(* IEC 61131-3 sources: trust-platform/examples/OSCAT/hvac_air_handling_unit/oop/src, 3 files *)

(* ---- Main.st ---- *)
(* Pattern role: IAhuStrategy is the contract boundary for the Strategy example. *)
INTERFACE IAhuStrategy EXTENDS IComponent
    PROPERTY ModeId : INT
    GET
    END_GET
    END_PROPERTY

    PROPERTY Output : REAL
    GET
    END_GET
    END_PROPERTY

    METHOD AcceptsCommand : BOOL
    VAR_INPUT
        SmokeClear : BOOL;
        FreezeStatClear : BOOL;
    END_VAR
    END_METHOD

    METHOD Update : REAL
    VAR_INPUT
        SupplyTemp : REAL;
        ScheduledSetpoint : REAL;
        OutdoorTemp : REAL;
    END_VAR
    END_METHOD
END_INTERFACE

(* Pattern role: EcoStrategy is a concrete implementation in the Strategy example. *)
FUNCTION_BLOCK EcoStrategy IMPLEMENTS IAhuStrategy
VAR
    ReadyValue : BOOL;
    ErrorValue : BOOL;
    ErrorIdValue : WORD;
    StatusValue : BYTE;
    OutputValue : REAL;
    Filter : Pt1Filter;
END_VAR

METHOD PUBLIC Initialize
ReadyValue := TRUE;
Filter.Initialize();
Filter.Configure(TimeConstant := T#5s, Gain := REAL#1.0);
ClearError();
END_METHOD

METHOD PUBLIC Reset
OutputValue := REAL#0.0;
ClearError();
END_METHOD

METHOD PUBLIC ClearError
ErrorValue := FALSE;
ErrorIdValue := WORD#0;
StatusValue := BYTE#0;
END_METHOD

METHOD PUBLIC Snapshot : ComponentStatus
VAR
    Result : ComponentStatus;
END_VAR
Result.Ready := ReadyValue;
Result.Error := ErrorValue;
Result.ErrorId := ErrorIdValue;
Result.Status := StatusValue;
Snapshot := Result;
END_METHOD

METHOD PUBLIC AcceptsCommand : BOOL
VAR_INPUT
    SmokeClear : BOOL;
    FreezeStatClear : BOOL;
END_VAR
AcceptsCommand := SmokeClear AND FreezeStatClear;
END_METHOD

METHOD PUBLIC Update : REAL
VAR_INPUT
    SupplyTemp : REAL;
    ScheduledSetpoint : REAL;
    OutdoorTemp : REAL;
END_VAR
VAR
    Error : REAL;
END_VAR
(* Filter is kept on the snapshot side for telemetry smoothing; the
   deadband and gain operate on the raw supply temp so the controller
   reacts to step changes within the same scan. *)
Filter.Update(Sample := SupplyTemp);
Error := ScheduledSetpoint - SupplyTemp;
IF ABS(Error) <= REAL#2.0 THEN
    OutputValue := REAL#0.0;
ELSE
    OutputValue := LIMIT(REAL#0.0, Error * REAL#8.0, REAL#100.0);
END_IF;
Update := OutputValue;
END_METHOD

PUBLIC PROPERTY ModeId : INT
GET
    ModeId := INT#1;
END_GET
END_PROPERTY

PUBLIC PROPERTY Output : REAL
GET
    Output := OutputValue;
END_GET
END_PROPERTY

PUBLIC PROPERTY Ready : BOOL
GET
    Ready := ReadyValue;
END_GET
END_PROPERTY

PUBLIC PROPERTY Error : BOOL
GET
    Error := ErrorValue;
END_GET
END_PROPERTY

PUBLIC PROPERTY ErrorId : WORD
GET
    ErrorId := ErrorIdValue;
END_GET
END_PROPERTY

PUBLIC PROPERTY Status : BYTE
GET
    Status := StatusValue;
END_GET
END_PROPERTY
END_FUNCTION_BLOCK

(* Pattern role: ComfortStrategy is a concrete implementation in the Strategy example. *)
FUNCTION_BLOCK ComfortStrategy IMPLEMENTS IAhuStrategy
VAR
    ReadyValue : BOOL;
    ErrorValue : BOOL;
    ErrorIdValue : WORD;
    StatusValue : BYTE;
    OutputValue : REAL;
    Filter : Pt1Filter;
END_VAR

METHOD PUBLIC Initialize
ReadyValue := TRUE;
Filter.Initialize();
Filter.Configure(TimeConstant := T#1s, Gain := REAL#1.0);
ClearError();
END_METHOD

METHOD PUBLIC Reset
OutputValue := REAL#0.0;
ClearError();
END_METHOD

METHOD PUBLIC ClearError
ErrorValue := FALSE;
ErrorIdValue := WORD#0;
StatusValue := BYTE#0;
END_METHOD

METHOD PUBLIC Snapshot : ComponentStatus
VAR
    Result : ComponentStatus;
END_VAR
Result.Ready := ReadyValue;
Result.Error := ErrorValue;
Result.ErrorId := ErrorIdValue;
Result.Status := StatusValue;
Snapshot := Result;
END_METHOD

METHOD PUBLIC AcceptsCommand : BOOL
VAR_INPUT
    SmokeClear : BOOL;
    FreezeStatClear : BOOL;
END_VAR
AcceptsCommand := SmokeClear;
END_METHOD

METHOD PUBLIC Update : REAL
VAR_INPUT
    SupplyTemp : REAL;
    ScheduledSetpoint : REAL;
    OutdoorTemp : REAL;
END_VAR
VAR
    Error : REAL;
END_VAR
(* Same approach as Eco: deadband/gain on raw supply, filter
   advanced for telemetry only. Strict inequality so Comfort reacts
   at the deadband boundary (tighter response than Eco). *)
Filter.Update(Sample := SupplyTemp);
Error := ScheduledSetpoint - SupplyTemp;
IF ABS(Error) < REAL#0.5 THEN
    OutputValue := REAL#0.0;
ELSE
    OutputValue := LIMIT(REAL#0.0, Error * REAL#20.0, REAL#100.0);
END_IF;
Update := OutputValue;
END_METHOD

PUBLIC PROPERTY ModeId : INT
GET
    ModeId := INT#2;
END_GET
END_PROPERTY

PUBLIC PROPERTY Output : REAL
GET
    Output := OutputValue;
END_GET
END_PROPERTY

PUBLIC PROPERTY Ready : BOOL
GET
    Ready := ReadyValue;
END_GET
END_PROPERTY

PUBLIC PROPERTY Error : BOOL
GET
    Error := ErrorValue;
END_GET
END_PROPERTY

PUBLIC PROPERTY ErrorId : WORD
GET
    ErrorId := ErrorIdValue;
END_GET
END_PROPERTY

PUBLIC PROPERTY Status : BYTE
GET
    Status := StatusValue;
END_GET
END_PROPERTY
END_FUNCTION_BLOCK

(* Pattern role: FrostProtectStrategy is a concrete implementation in the Strategy example. *)
FUNCTION_BLOCK FrostProtectStrategy IMPLEMENTS IAhuStrategy
VAR
    ReadyValue : BOOL;
    ErrorValue : BOOL;
    ErrorIdValue : WORD;
    StatusValue : BYTE;
    OutputValue : REAL;
END_VAR

METHOD PUBLIC Initialize
ReadyValue := TRUE;
ClearError();
END_METHOD

METHOD PUBLIC Reset
OutputValue := REAL#0.0;
ClearError();
END_METHOD

METHOD PUBLIC ClearError
ErrorValue := FALSE;
ErrorIdValue := WORD#0;
StatusValue := BYTE#0;
END_METHOD

METHOD PUBLIC Snapshot : ComponentStatus
VAR
    Result : ComponentStatus;
END_VAR
Result.Ready := ReadyValue;
Result.Error := ErrorValue;
Result.ErrorId := ErrorIdValue;
Result.Status := StatusValue;
Snapshot := Result;
END_METHOD

METHOD PUBLIC AcceptsCommand : BOOL
VAR_INPUT
    SmokeClear : BOOL;
    FreezeStatClear : BOOL;
END_VAR
AcceptsCommand := SmokeClear;
END_METHOD

METHOD PUBLIC Update : REAL
VAR_INPUT
    SupplyTemp : REAL;
    ScheduledSetpoint : REAL;
    OutdoorTemp : REAL;
END_VAR
VAR
    FrostTarget : REAL;
END_VAR
FrostTarget := MAX(ScheduledSetpoint, REAL#5.0);
OutputValue := LIMIT(REAL#20.0, (FrostTarget - SupplyTemp) * REAL#30.0, REAL#100.0);
Update := OutputValue;
END_METHOD

PUBLIC PROPERTY ModeId : INT
GET
    ModeId := INT#3;
END_GET
END_PROPERTY

PUBLIC PROPERTY Output : REAL
GET
    Output := OutputValue;
END_GET
END_PROPERTY

PUBLIC PROPERTY Ready : BOOL
GET
    Ready := ReadyValue;
END_GET
END_PROPERTY

PUBLIC PROPERTY Error : BOOL
GET
    Error := ErrorValue;
END_GET
END_PROPERTY

PUBLIC PROPERTY ErrorId : WORD
GET
    ErrorId := ErrorIdValue;
END_GET
END_PROPERTY

PUBLIC PROPERTY Status : BYTE
GET
    Status := StatusValue;
END_GET
END_PROPERTY
END_FUNCTION_BLOCK

(* Composition role: AhuController owns the collaborating objects used by this Strategy example. *)
FUNCTION_BLOCK AhuController
VAR
    Eco : EcoStrategy;
    Comfort : ComfortStrategy;
    Frost : FrostProtectStrategy;
    ActiveStrategy : IAhuStrategy;
    StateValue : INT;
    ActiveModeValue : INT;
    HeatingCommandValue : REAL;
    AlarmActiveValue : BOOL;
    AlarmCodeValue : DWORD;
    RuntimeFan : OntimeMeter;
    AlarmQueue : DwordFifo16;
END_VAR

METHOD PUBLIC Initialize
Eco.Initialize();
Comfort.Initialize();
Frost.Initialize();
RuntimeFan.Initialize();
RuntimeFan.Reset();
AlarmQueue.Initialize();
AlarmQueue.Reset();
StateValue := INT#0;
ActiveModeValue := INT#0;
HeatingCommandValue := REAL#0.0;
AlarmActiveValue := FALSE;
AlarmCodeValue := DWORD#0;
END_METHOD

METHOD PRIVATE RaiseAlarm
VAR_INPUT
    Code : DWORD;
END_VAR
AlarmActiveValue := TRUE;
AlarmCodeValue := Code;
StateValue := INT#900;
IF AlarmQueue.Push(Value := Code) THEN
END_IF;
END_METHOD

METHOD PUBLIC Update : REAL
VAR_INPUT
    ModeRequest : INT;
    OutdoorTemp : REAL;
    SupplyTemp : REAL;
    SupplySetpoint : REAL;
    SmokeClear : BOOL;
    FreezeStatClear : BOOL;
    SupplyFanHealthy : BOOL;
END_VAR
IF NOT SmokeClear THEN
    RaiseAlarm(Code := DWORD#16#A100);
    HeatingCommandValue := REAL#0.0;
ELSE
    IF (OutdoorTemp < REAL#-5.0) OR NOT FreezeStatClear THEN
        ActiveStrategy := Frost;
    ELSIF ModeRequest = INT#1 THEN
        ActiveStrategy := Eco;
    ELSE
        ActiveStrategy := Comfort;
    END_IF;

    ActiveModeValue := ActiveStrategy.ModeId;
    IF NOT SupplyFanHealthy THEN
        RaiseAlarm(Code := DWORD#16#A101);
    ELSIF ActiveStrategy.AcceptsCommand(SmokeClear := SmokeClear, FreezeStatClear := FreezeStatClear) THEN
        StateValue := INT#200;
        HeatingCommandValue := ActiveStrategy.Update(SupplyTemp := SupplyTemp, ScheduledSetpoint := SupplySetpoint, OutdoorTemp := OutdoorTemp);
        RuntimeFan.Update(Input := TRUE);
    ELSE
        RaiseAlarm(Code := DWORD#16#B100);
    END_IF;
END_IF;
Update := HeatingCommandValue;
END_METHOD

PUBLIC PROPERTY State : INT
GET
    State := StateValue;
END_GET
END_PROPERTY

PUBLIC PROPERTY ActiveMode : INT
GET
    ActiveMode := ActiveModeValue;
END_GET
END_PROPERTY

PUBLIC PROPERTY HeatingCommand : REAL
GET
    HeatingCommand := HeatingCommandValue;
END_GET
END_PROPERTY

PUBLIC PROPERTY AlarmActive : BOOL
GET
    AlarmActive := AlarmActiveValue;
END_GET
END_PROPERTY
END_FUNCTION_BLOCK

(* Scan role: Main wires the example objects and exposes the PLC call path under test. *)
PROGRAM Main
VAR
    Ahu : AhuController;
    Initialized : BOOL;
    ModeRequest : INT;
    OutdoorTempRaw : INT;
    SupplyTempRaw : INT;
    SmokeClear : BOOL;
    FreezeStatClear : BOOL;
    SupplyFanHealthy : BOOL;
    HeatingValveRaw : INT;
    SupplyFanEnable : BOOL;
    FireAlarmRelay : BOOL;
    OutdoorTemp : REAL;
    SupplyTemp : REAL;
END_VAR

OutdoorTemp := TO_REAL(OutdoorTempRaw) / REAL#10.0;
SupplyTemp := TO_REAL(SupplyTempRaw) / REAL#10.0;
(* Initialize once on cold start; scanning Initialize every cycle would
   reset RuntimeFan, clear AlarmQueue, and force StateValue back to 0. *)
IF NOT Initialized THEN
    Ahu.Initialize();
    Initialized := TRUE;
END_IF;
HeatingValveRaw := TO_INT(Ahu.Update(ModeRequest := ModeRequest, OutdoorTemp := OutdoorTemp, SupplyTemp := SupplyTemp, SupplySetpoint := REAL#21.0, SmokeClear := SmokeClear, FreezeStatClear := FreezeStatClear, SupplyFanHealthy := SupplyFanHealthy) * REAL#10.0);
SupplyFanEnable := NOT Ahu.AlarmActive;
FireAlarmRelay := NOT SmokeClear;
END_PROGRAM

(* ---- Configuration.st ---- *)
CONFIGURATION AhuOopConfiguration
RESOURCE AhuOop ON PLC
    TASK MainTask (INTERVAL := T#100ms, PRIORITY := 1);
    PROGRAM Ahu WITH MainTask : Main;
END_RESOURCE
VAR_CONFIG
    Ahu.ModeRequest AT %IW0 : INT;
    Ahu.OutdoorTempRaw AT %IW2 : INT;
    Ahu.SupplyTempRaw AT %IW4 : INT;
    Ahu.SmokeClear AT %IX0.0 : BOOL;
    Ahu.FreezeStatClear AT %IX0.1 : BOOL;
    Ahu.SupplyFanHealthy AT %IX0.2 : BOOL;
    Ahu.HeatingValveRaw AT %QW0 : INT;
    Ahu.SupplyFanEnable AT %QX0.0 : BOOL;
    Ahu.FireAlarmRelay AT %QX0.1 : BOOL;
END_VAR
END_CONFIGURATION

(* ---- Tests.st ---- *)
TEST_PROGRAM AhuStrategySelectsModeSpecificObjects
VAR
    Ahu : AhuController;
    EcoCommand : REAL;
    ComfortCommand : REAL;
    FrostCommand : REAL;
END_VAR

Ahu.Initialize();
EcoCommand := Ahu.Update(ModeRequest := INT#1, OutdoorTemp := REAL#10.0, SupplyTemp := REAL#18.0, SupplySetpoint := REAL#21.0, SmokeClear := TRUE, FreezeStatClear := TRUE, SupplyFanHealthy := TRUE);
ASSERT_EQUAL(EXPECTED := INT#1, ACTUAL := Ahu.ActiveMode);

ComfortCommand := Ahu.Update(ModeRequest := INT#2, OutdoorTemp := REAL#10.0, SupplyTemp := REAL#18.0, SupplySetpoint := REAL#21.0, SmokeClear := TRUE, FreezeStatClear := TRUE, SupplyFanHealthy := TRUE);
ASSERT_EQUAL(EXPECTED := INT#2, ACTUAL := Ahu.ActiveMode);
ASSERT_TRUE(IN := ComfortCommand > EcoCommand);

FrostCommand := Ahu.Update(ModeRequest := INT#1, OutdoorTemp := REAL#-8.0, SupplyTemp := REAL#1.0, SupplySetpoint := REAL#3.0, SmokeClear := TRUE, FreezeStatClear := FALSE, SupplyFanHealthy := TRUE);
ASSERT_EQUAL(EXPECTED := INT#3, ACTUAL := Ahu.ActiveMode);
ASSERT_TRUE(IN := FrostCommand >= REAL#20.0);
END_TEST_PROGRAM

TEST_PROGRAM AhuSmokeAlarmOverridesAllStrategies
VAR
    Ahu : AhuController;
    Command : REAL;
END_VAR

Ahu.Initialize();
Command := Ahu.Update(ModeRequest := INT#2, OutdoorTemp := REAL#10.0, SupplyTemp := REAL#18.0, SupplySetpoint := REAL#21.0, SmokeClear := FALSE, FreezeStatClear := TRUE, SupplyFanHealthy := TRUE);
ASSERT_TRUE(IN := Ahu.AlarmActive);
ASSERT_NEAR(EXPECTED := REAL#0.0, ACTUAL := Command, DELTA := REAL#0.001);
END_TEST_PROGRAM

(* Integration test: simulates the PROGRAM Main scan loop with the
   Init-once guard. Catches the "Initialize every cycle" bug —
   AhuController.Initialize() resets RuntimeFan accumulator, clears
   AlarmQueue, and forces State back to 0. Without the guard, the
   active mode never persists across cycles. *)
TEST_PROGRAM AhuScanLoopWithInitGuardPersistsActiveModeAcrossCycles
VAR
    Ahu : AhuController;
    Initialized : BOOL;
    I : INT;
    LastMode : INT;
END_VAR

FOR I := 1 TO 5 DO
    IF NOT Initialized THEN
        Ahu.Initialize();
        Initialized := TRUE;
    END_IF;
    Ahu.Update(ModeRequest := INT#2, OutdoorTemp := REAL#10.0, SupplyTemp := REAL#18.0, SupplySetpoint := REAL#21.0, SmokeClear := TRUE, FreezeStatClear := TRUE, SupplyFanHealthy := TRUE);
    LastMode := Ahu.ActiveMode;
END_FOR;
(* After five cycles in Comfort mode, the active mode is stable *)
ASSERT_EQUAL(EXPECTED := INT#2, ACTUAL := LastMode);
ASSERT_FALSE(IN := Ahu.AlarmActive);
END_TEST_PROGRAM

(* Anti-pattern test: re-initializing every cycle resets all retained
   state. This pins the contract: if a future change removes the
   Init-once guard from Main, this test still passes (because the
   anti-pattern is what's tested), but the guard test above will fail
   if the assertion is ever violated by re-init mid-flight. *)
TEST_PROGRAM AhuReinitializingEveryCycleClearsAlarmsAndState
VAR
    Ahu : AhuController;
    I : INT;
END_VAR

(* Trip a smoke alarm, then re-init: alarm should clear *)
Ahu.Initialize();
Ahu.Update(ModeRequest := INT#2, OutdoorTemp := REAL#10.0, SupplyTemp := REAL#18.0, SupplySetpoint := REAL#21.0, SmokeClear := FALSE, FreezeStatClear := TRUE, SupplyFanHealthy := TRUE);
ASSERT_TRUE(IN := Ahu.AlarmActive);
Ahu.Initialize();
ASSERT_FALSE(IN := Ahu.AlarmActive);
END_TEST_PROGRAM

(* FrostProtect override priority: outdoor < -5 forces Frost regardless of mode request. *)
TEST_PROGRAM AhuFrostProtectOverridesAllOtherModes
VAR
    Ahu : AhuController;
END_VAR
Ahu.Initialize();

(* Eco request but freezing outside - Frost wins *)
Ahu.Update(ModeRequest := INT#1, OutdoorTemp := REAL#-10.0, SupplyTemp := REAL#5.0, SupplySetpoint := REAL#21.0, SmokeClear := TRUE, FreezeStatClear := TRUE, SupplyFanHealthy := TRUE);
ASSERT_EQUAL(EXPECTED := INT#3, ACTUAL := Ahu.ActiveMode);

(* Comfort request but freezing - Frost wins *)
Ahu.Update(ModeRequest := INT#2, OutdoorTemp := REAL#-10.0, SupplyTemp := REAL#5.0, SupplySetpoint := REAL#21.0, SmokeClear := TRUE, FreezeStatClear := TRUE, SupplyFanHealthy := TRUE);
ASSERT_EQUAL(EXPECTED := INT#3, ACTUAL := Ahu.ActiveMode);

(* Boundary: outdoor exactly -5 (NOT below -5, strict less-than) - Eco wins *)
Ahu.Update(ModeRequest := INT#1, OutdoorTemp := REAL#-5.0, SupplyTemp := REAL#15.0, SupplySetpoint := REAL#21.0, SmokeClear := TRUE, FreezeStatClear := TRUE, SupplyFanHealthy := TRUE);
ASSERT_EQUAL(EXPECTED := INT#1, ACTUAL := Ahu.ActiveMode);

(* Freeze stat trip alone (warm outside) -> Frost still wins *)
Ahu.Update(ModeRequest := INT#1, OutdoorTemp := REAL#15.0, SupplyTemp := REAL#15.0, SupplySetpoint := REAL#21.0, SmokeClear := TRUE, FreezeStatClear := FALSE, SupplyFanHealthy := TRUE);
ASSERT_EQUAL(EXPECTED := INT#3, ACTUAL := Ahu.ActiveMode);
END_TEST_PROGRAM

(* Smoke is the highest priority - it wins over Frost. *)
TEST_PROGRAM AhuSmokeBeatsFrostProtect
VAR
    Ahu : AhuController;
    Command : REAL;
END_VAR
Ahu.Initialize();

(* Both smoke and freeze conditions present -> alarm + heat off *)
Command := Ahu.Update(ModeRequest := INT#1, OutdoorTemp := REAL#-10.0, SupplyTemp := REAL#0.0, SupplySetpoint := REAL#5.0, SmokeClear := FALSE, FreezeStatClear := FALSE, SupplyFanHealthy := TRUE);
ASSERT_TRUE(IN := Ahu.AlarmActive);
ASSERT_NEAR(EXPECTED := REAL#0.0, ACTUAL := Command, DELTA := REAL#0.001);
END_TEST_PROGRAM

(* Eco strategy: deadband of +/- 2 C around setpoint. *)
TEST_PROGRAM AhuEcoStrategyHasWideDeadband
VAR
    Eco : EcoStrategy;
    Out : REAL;
END_VAR
Eco.Initialize();

(* Inside +/- 2 C deadband -> output 0 *)
Out := Eco.Update(SupplyTemp := REAL#21.0, ScheduledSetpoint := REAL#21.0, OutdoorTemp := REAL#10.0);
ASSERT_NEAR(EXPECTED := REAL#0.0, ACTUAL := Out, DELTA := REAL#0.001);

Out := Eco.Update(SupplyTemp := REAL#19.5, ScheduledSetpoint := REAL#21.0, OutdoorTemp := REAL#10.0);
ASSERT_NEAR(EXPECTED := REAL#0.0, ACTUAL := Out, DELTA := REAL#0.001);

(* Outside deadband -> non-zero command *)
Out := Eco.Update(SupplyTemp := REAL#15.0, ScheduledSetpoint := REAL#21.0, OutdoorTemp := REAL#10.0);
ASSERT_TRUE(IN := Out > REAL#0.0);
END_TEST_PROGRAM

(* Comfort strategy: tighter deadband (+/- 0.5 C) and higher gain. *)
TEST_PROGRAM AhuComfortStrategyTighterThanEco
VAR
    Comfort : ComfortStrategy;
    Eco : EcoStrategy;
    ComfortOut : REAL;
    EcoOut : REAL;
END_VAR
Comfort.Initialize();
Eco.Initialize();

(* Same input - Comfort produces higher output (gain 20 vs Eco's 8) *)
ComfortOut := Comfort.Update(SupplyTemp := REAL#19.0, ScheduledSetpoint := REAL#21.0, OutdoorTemp := REAL#10.0);
EcoOut := Eco.Update(SupplyTemp := REAL#19.0, ScheduledSetpoint := REAL#21.0, OutdoorTemp := REAL#10.0);
ASSERT_TRUE(IN := ComfortOut > EcoOut);

(* Comfort responds to small errors that Eco ignores *)
ComfortOut := Comfort.Update(SupplyTemp := REAL#20.5, ScheduledSetpoint := REAL#21.0, OutdoorTemp := REAL#10.0);
EcoOut := Eco.Update(SupplyTemp := REAL#20.5, ScheduledSetpoint := REAL#21.0, OutdoorTemp := REAL#10.0);
ASSERT_NEAR(EXPECTED := REAL#0.0, ACTUAL := EcoOut, DELTA := REAL#0.001);
ASSERT_TRUE(IN := ComfortOut > REAL#0.0);
END_TEST_PROGRAM

(* FrostProtect strategy: forces setpoint to MAX(scheduled, 5 C). *)
TEST_PROGRAM AhuFrostProtectClampsSetpointToMinimumFiveCelsius
VAR
    Frost : FrostProtectStrategy;
    Out : REAL;
END_VAR
Frost.Initialize();

(* Scheduled setpoint below 5 C - Frost forces to 5 *)
Out := Frost.Update(SupplyTemp := REAL#3.0, ScheduledSetpoint := REAL#0.0, OutdoorTemp := REAL#-10.0);
(* Effective setpoint 5, error 2, gain 30 -> output ~60, then LIMITed to 100 max but at least 20 min *)
ASSERT_TRUE(IN := Out >= REAL#20.0);

(* Scheduled setpoint above 5 - Frost uses scheduled *)
Out := Frost.Update(SupplyTemp := REAL#15.0, ScheduledSetpoint := REAL#21.0, OutdoorTemp := REAL#-10.0);
ASSERT_TRUE(IN := Out > REAL#0.0);

(* Output never falls below 20 even when error is small (forced minimum heat) *)
Out := Frost.Update(SupplyTemp := REAL#21.0, ScheduledSetpoint := REAL#21.0, OutdoorTemp := REAL#-10.0);
ASSERT_TRUE(IN := Out >= REAL#20.0);
END_TEST_PROGRAM

(* Supply fan unhealthy raises a class B alarm. *)
TEST_PROGRAM AhuSupplyFanFaultRaisesAlarm
VAR
    Ahu : AhuController;
END_VAR
Ahu.Initialize();
Ahu.Update(ModeRequest := INT#2, OutdoorTemp := REAL#10.0, SupplyTemp := REAL#18.0, SupplySetpoint := REAL#21.0, SmokeClear := TRUE, FreezeStatClear := TRUE, SupplyFanHealthy := FALSE);
ASSERT_TRUE(IN := Ahu.AlarmActive);
END_TEST_PROGRAM
